(* IEC 61131-3 sources: Caravan/Archiv/12-04-19/Stations/Terminal/HMI/Network/LseRtkMain, 1 file *)

(* ---- ONE_LseRtkMain_Table.st ---- *)
#define OBJECTS_CONFIG

FUNCTION GLOBAL TAB ONE_LseRtkMain
-1$UINT, 0$UINT,
0$UINT, 0$UINT,

3$UDINT,
TO_UDINT(1552551876), "_Lse", 0$UINT, 114$UINT, 1$UINT,
TO_UDINT(3931827689), "_SysDateTime", 0$UINT, 7$UINT, 1$UINT,
TO_UDINT(1903583397), "Ram", 1$UINT, 3$UINT, 1$UINT,

_NO_ATTR, TO_UDINT(299963966), "LSE",

_NO_ATTR, TO_UDINT(3035062039), "SYSDATETIME",

1$UINT, TO_UDINT(1119588755), "SYSDATETIME\SUMMERTIME",

//Internal connections
0$UDINT,
1$UDINT,
TO_UDINT(1), "SummerTime", TO_UDINT(2),
0$UDINT,
0$UDINT,

//Initialization values
0$UDINT,
3$UDINT,
TO_UDINT(0), "AmericanDateFormat", TO_UDINT(0),//|LseRtkMain.Lse.AmericanDateFormat;
TO_UDINT(0), "SeekAlgorithm", TO_UDINT(1),//|LseRtkMain.Lse.SeekAlgorithm;
TO_UDINT(1), "DoSummerTime", TO_UDINT(0),//|LseRtkMain.SysDateTime.DoSummerTime;

//Symbolic initialization values
0$UDINT,
0$UDINT,

//Initialization of string values
0$UDINT,
0$UDINT,

//Configuration of tasks (RealTime, Cyclic, Background)
0$UDINT,
0$UDINT,

0$UDINT,
0$UDINT,

0$UDINT,
2$UDINT,
TO_UDINT(0), (-1)$UDINT, 4194303$DINT, 	//LSE
TO_UDINT(1), (100)$UDINT, 4194303$DINT, 	//SYSDATETIME

//External connections
0$UDINT,
0$UDINT,

//Magic internal connections
0$UDINT,
0$UDINT,

//Configuration of timeslots of tasks (RealTime, Cyclic)
#ifdef __LSLLDR_TIMESLOTS__
0$UDINT,
0$UDINT,

0$UDINT,
0$UDINT,

#endif //__LSLLDR_TIMESLOTS__

//MultiMaster connections
#ifdef __LSLLDR_MULTIMASTER__
0$UDINT,
0$UDINT,
#endif //__LSLLDR_MULTIMASTER__

//Configuration for task ID (RealTime, CyclicTime)
#ifdef __LSLLDR_TASKID__
"\\\\TASKS2  "
0$UDINT,
0$UDINT,

0$UDINT,
0$UDINT,

0$UDINT,
2$UDINT,
(0)$UDINT, 	//LSE
(0)$UDINT, 	//SYSDATETIME

#endif //__LSLLDR_TASKID__

END_FUNCTION
